                                   //LCom Version V1
                                   #statSend.tsendFct.data[#statSend.tsendFct.dataOffset] := #statSend.configTelegramV1.LComVersion;
                                   #statSend.tsendFct.data[#statSend.tsendFct.dataOffset + 1] := 16#03;
                                   #statSend.tsendFct.data[#statSend.tsendFct.dataOffset + 2] := #statSend.configTelegramV1.comMode;//ComMode
                                   #statSend.tsendFct.data[#statSend.tsendFct.dataOffset + 3] := #statSend.configTelegramV1.slidingWindow;//SlidingWindow
                                   //cycleTime
                                   #statSend.tsendFct.data[#statSend.tsendFct.dataOffset + 4] := #statSend.configTelegramV1.cycleTime.%B1;
                                   #statSend.tsendFct.data[#statSend.tsendFct.dataOffset + 5] := #statSend.configTelegramV1.cycleTime.%B0;
                                   //ackTimeOut
                                   #statSend.tsendFct.data[#statSend.tsendFct.dataOffset + 6] := #statSend.configTelegramV1.ackTimeOut.%B1;
                                   #statSend.tsendFct.data[#statSend.tsendFct.dataOffset + 7] := #statSend.configTelegramV1.ackTimeOut.%B0;
                                   //lifeSignCycle
                                   #statSend.tsendFct.data[#statSend.tsendFct.dataOffset + 8] := #statSend.configTelegramV1.lifeSignCycle.%B1;
                                   #statSend.tsendFct.data[#statSend.tsendFct.dataOffset + 9] := #statSend.configTelegramV1.lifeSignCycle.%B0;
                                   //status
                                   #statSend.tsendFct.data[#statSend.tsendFct.dataOffset + 10] := #statSend.configTelegramV1.status;
                                   //sendModeSyncTime
                                   #statSend.tsendFct.data[#statSend.tsendFct.dataOffset + 11] := #statSend.configTelegramV1.sendModeSyncTime;
                                   //maxSendDataLength
                                   #statSend.tsendFct.data[#statSend.tsendFct.dataOffset + 12] := #statSend.configTelegramV1.maxSendDataLength.%B1;
                                   #statSend.tsendFct.data[#statSend.tsendFct.dataOffset + 13] := #statSend.configTelegramV1.maxSendDataLength.%B0;
                                   //maxReceiveDataLength
                                   #statSend.tsendFct.data[#statSend.tsendFct.dataOffset + 14] := #statSend.configTelegramV1.maxReceiveDataLength.%B1;
                                   #statSend.tsendFct.data[#statSend.tsendFct.dataOffset + 15] := #statSend.configTelegramV1.maxReceiveDataLength.%B0;
                                   //calculate new offset
                                   #statSend.tsendFct.dataOffset := 16;
                               ELSE
                                   #statSend.tsendFct.data[#statSend.tsendFct.dataOffset] := #statSend.configTelegramV2.LComVersion;
                                   #statSend.tsendFct.data[#statSend.tsendFct.dataOffset + 1] := 16#03;
                                   //status
                                   #statSend.tsendFct.data[#statSend.tsendFct.dataOffset + 2] := #statSend.configTelegramV2.status;
                                   //sendModeSyncTime
                                   #statSend.tsendFct.data[#statSend.tsendFct.dataOffset + 3] := #statSend.configTelegramV2.sendModeSyncTime;
                                   //lifeSignCycle
                                   #tempDWord := TIME_TO_DWORD(#statSend.configTelegramV2.lifeSignCycle);
                                   #statSend.tsendFct.data[#statSend.tsendFct.dataOffset + 4] := #tempDWord.%B3;
                                   #statSend.tsendFct.data[#statSend.tsendFct.dataOffset + 5] := #tempDWord.%B2;
                                   #statSend.tsendFct.data[#statSend.tsendFct.dataOffset + 6] := #tempDWord.%B1;
                                   #statSend.tsendFct.data[#statSend.tsendFct.dataOffset + 7] := #tempDWord.%B0;
                                   //cycleTime
                                   #tempDWord := TIME_TO_DWORD(#statSend.configTelegramV2.cycleTime);
                                   #statSend.tsendFct.data[#statSend.tsendFct.dataOffset + 8] := #tempDWord.%B3;
                                   #statSend.tsendFct.data[#statSend.tsendFct.dataOffset + 9] := #tempDWord.%B2;
                                   #statSend.tsendFct.data[#statSend.tsendFct.dataOffset + 10] := #tempDWord.%B1;
                                   #statSend.tsendFct.data[#statSend.tsendFct.dataOffset + 11] := #tempDWord.%B0;
                                   //ackTimeOut
                                   #tempDWord := TIME_TO_DWORD(#statSend.configTelegramV2.ackTimeOut);
                                   #statSend.tsendFct.data[#statSend.tsendFct.dataOffset + 12] := #tempDWord.%B3;
                                   #statSend.tsendFct.data[#statSend.tsendFct.dataOffset + 13] := #tempDWord.%B2;
                                   #statSend.tsendFct.data[#statSend.tsendFct.dataOffset + 14] := #tempDWord.%B1;
                                   #statSend.tsendFct.data[#statSend.tsendFct.dataOffset + 15] := #tempDWord.%B0;
                                   //maxSendDataLength
                                   #statSend.tsendFct.data[#statSend.tsendFct.dataOffset + 16] := #statSend.configTelegramV2.maxSendDataLength.%B3;
                                   #statSend.tsendFct.data[#statSend.tsendFct.dataOffset + 17] := #statSend.configTelegramV2.maxSendDataLength.%B2;
                                   #statSend.tsendFct.data[#statSend.tsendFct.dataOffset + 18] := #statSend.configTelegramV2.maxSendDataLength.%B1;
                                   #statSend.tsendFct.data[#statSend.tsendFct.dataOffset + 19] := #statSend.configTelegramV2.maxSendDataLength.%B0;
                                   //maxReceiveDataLength
                                   #statSend.tsendFct.data[#statSend.tsendFct.dataOffset + 20] := #statSend.configTelegramV2.maxReceiveDataLength.%B3;
                                   #statSend.tsendFct.data[#statSend.tsendFct.dataOffset + 21] := #statSend.configTelegramV2.maxReceiveDataLength.%B2;
                                   #statSend.tsendFct.data[#statSend.tsendFct.dataOffset + 22] := #statSend.configTelegramV2.maxReceiveDataLength.%B1;
                                   #statSend.tsendFct.data[#statSend.tsendFct.dataOffset + 23] := #statSend.configTelegramV2.maxReceiveDataLength.%B0;
                                   //calculate new offset
                                   #statSend.tsendFct.dataOffset := 24;
                               END_IF;
                               #statSend.tsendFct.enable := TRUE;

                               #instLocalLifeSignCycleTimer(IN := FALSE,
                                                            PT := #diagnostics.localConfig.connection.lifeSignCycleTime);
                           ELSE
                               ;//Telegram 3 don´t need be send

                           END_IF;
                       ELSIF (NOT #diagnostics.localConfig.connection.useLComProtocol //without LCom Protocol
                           AND #statState.sender = #STATE_INACTIVE) THEN
                           #statSend.tsendFct.enable := FALSE;
                       ELSE
                           #statSend.tsendFct.enable := TRUE;

                           #instLocalLifeSignCycleTimer(IN := FALSE,
                                                        PT := #diagnostics.localConfig.connection.lifeSignCycleTime);
                       END_IF;

                       //differ between different connection types (IPv4, QDN)
                       IF (#diagnostics.localConfig.connection.connectType = #CON_TYPE_IPV4) THEN
                           #tempConnOucId := #statTconPar.ID;
                       ELSE    //#CON_TYPE_QDN
                           #tempConnOucId := #statTconParQdn.ID;
                       END_IF;

                       #instTSEND(REQ := #statSend.tsendFct.enable,
                                  LEN := #statSend.tsendFct.dataOffset,
                                  ID := #tempConnOucId,
                                  DATA := #statSend.tsendFct.data,
                                  STATUS => #statSend.tsendFct.status);

                       //16#80C4=Temporary communication error
                       IF (#statSend.tsendFct.status = 16#80C4) THEN

                           #instSendErrorTimer(IN := TRUE,
                                               PT := #MAX_TRIAL_TIME);

                           //#MAX_TRIAL_TIME is expired
                           IF #instSendErrorTimer.Q THEN
                               //Write diagnostics
                               #statDiag.bufferIndex := #statDiag.bufferIndex + 1;
                               #statDiag.buffer[#statDiag.bufferIndex].status := #ERR_SEND;
                               #statDiag.buffer[#statDiag.bufferIndex].subFunctionErrorID := #statSend.tsendFct.status;
                               #statDiag.buffer[#statDiag.bufferIndex].additionalValue1 := 0.0;
                               #statDiag.buffer[#statDiag.bufferIndex].additionalValue2 := #statSend.tsendFct.dataOffset;
                               #statDiag.buffer[#statDiag.bufferIndex].additionalValue3 := 0.0;
                               #statDiag.buffer[#statDiag.bufferIndex].additionalValue4 := T#0ms;
                               #statState.connection := #CLOSE_CONNECTION;
                               GOTO diag;
                           END_IF;
                       ELSIF (#statSend.tsendFct.status >= 16#8085) THEN
                           //#WARN_SEND
                           #statDiag.bufferIndex := #statDiag.bufferIndex + 1;
                           #statDiag.buffer[#statDiag.bufferIndex].status := #ERR_SEND;
                           #statDiag.buffer[#statDiag.bufferIndex].subFunctionErrorID := #statSend.tsendFct.status;
                           #statDiag.buffer[#statDiag.bufferIndex].additionalValue1 := 0.0;
                           #statDiag.buffer[#statDiag.bufferIndex].additionalValue2 := #statSend.tsendFct.dataOffset;
                           #statDiag.buffer[#statDiag.bufferIndex].additionalValue3 := 0.0;
                           #statDiag.buffer[#statDiag.bufferIndex].additionalValue4 := T#0ms;

                           #statState.connection := #CLOSE_CONNECTION;
                           GOTO diag;
                       END_IF;
                   END_REGION SEND_LIFESIGN

               END_REGION OPERATION

           #STATE_INACTIVE_PREPARE:
               REGION INACTIVE_PREPARE

                   #statState.connection := #STATE_INACTIVE;
                   #status := #statStatus := #STATUS_NO_CALL;
                   #statFallingEdgeEnable := FALSE;
                   #statOldEnable := FALSE;
                   #busy := FALSE;
               END_REGION INACTIVE_PREPARE

           #STATE_INIT:
               REGION INIT
                   //Reset FB Outputs
                   #connected := #statConnected := FALSE;
                   #sending := #statSending := FALSE;
                   #error := FALSE;

                   //Diagnostics purpose
                   //connection
                   #diagnostics.localConfig.connection.connectionID := #configuration.connection.connectionID;
                   #diagnostics.localConfig.connection.interfaceID := #configuration.connection.interfaceID;
                   #diagnostics.localConfig.connection.comService := #configuration.connection.comService;
                   #diagnostics.localConfig.connection.isClient := #configuration.connection.isClient;
                   #diagnostics.localConfig.connection.localPort := #configuration.connection.localPort;
                   #diagnostics.localConfig.connection.partnerPort := #configuration.connection.partnerPort;
                   #diagnostics.localConfig.connection.partnerIP := #configuration.connection.partnerIP;
                   #diagnostics.localConfig.connection.acceptUnknownPartner := #configuration.connection.acceptUnknownPartner;
                   #statActualLocalLComVersion := #HEADER_V2;
                   #diagnostics.localConfig.connection.lifeSignCycleTime := #configuration.connection.lifeSignCycleTime;
                   //-->QDN
                   #diagnostics.localConfig.connection.connectType := #configuration.connection.connectType;
                   #diagnostics.localConfig.connection.partnerQDN := #configuration.connection.partnerQDN;
                   //Sender
                   #diagnostics.localConfig.sender.cycleTime := #configuration.sender.cycleTime;
                   #diagnostics.localConfig.sender.ackTimeout := #configuration.sender.ackTimeout;
                   //TimeSync
                   #diagnostics.localConfig.timeSync.usePartnerTimestamps := #configuration.timeSync.usePartnerTimestamps;
                   #diagnostics.localConfig.timeSync.sendMode := #configuration.timeSync.sendMode;
                   #diagnostics.localConfig.timeSync.cycleTime := #configuration.timeSync.cycleTime;
                   #diagnostics.localConfig.timeSync.sendAtTimeOfDay := #configuration.timeSync.sendAtTimeOfDay;
                   //Statistics
                   #diagnostics.statistics.avgCallCycle := 0.0;
                   #diagnostics.statistics.avgReceiveMsgCycle := 0.0;
                   #diagnostics.statistics.maxReceiveMsgCycle := T#0ms;
                   #diagnostics.statistics.LComProtocolUsed := FALSE;
                   #diagnostics.statistics.activeLComVersion := 0;
                   #diagnostics.statistics.avgMsgSendingTime := 0.0;
                   #diagnostics.statistics.maxMsgSendingTime := T#0ms;
                   #diagnostics.statistics.avgMsgReceivingTime := 0.0;
                   #diagnostics.statistics.maxMsgReceivingTime := T#0ms;
                   #diagnostics.statistics.numberOfSentMessages := 0;
                   #diagnostics.statistics.numberOfReceivedMessages := 0;
                   #diagnostics.statistics.totalAckTimeouts := 0;
                   #diagnostics.statistics.totalSendCycleViolations := 0;
                   #diagnostics.statistics.totalReceiveCycleViolations := 0;
                   #diagnostics.statistics.totalReconnects := 0;

                   #statConnectAttempts := 0;

                   //Check hardware identifier of the local interface
                   IF ((#diagnostics.localConfig.connection.interfaceID >= 0) //(0...65535)
                       AND
                       (#diagnostics.localConfig.connection.interfaceID <= 65535))
                   THEN
                       //Hardware identifier of the local interface --> OK
                       #statTconPar.InterfaceId := #diagnostics.localConfig.connection.interfaceID;
                   ELSE
                       //Hardware identifier of the local interface --> NOT OK
                       #statDiag.bufferIndex := #statDiag.bufferIndex + 1;
                       #statDiag.buffer[#statDiag.bufferIndex].status := #ERR_INTERFACE_ID;
                       #statDiag.buffer[#statDiag.bufferIndex].subFunctionErrorID := 16#0000;
                       #statDiag.buffer[#statDiag.bufferIndex].additionalValue1 := UINT_TO_REAL(#diagnostics.localConfig.connection.interfaceID);//value from user
                       #statDiag.buffer[#statDiag.bufferIndex].additionalValue2 := 0.0;
                       #statDiag.buffer[#statDiag.bufferIndex].additionalValue3 := 0.0;
                       #statDiag.buffer[#statDiag.bufferIndex].additionalValue4 := T#0ms;

                       #statState.connection := #ERROR_STATE;
                       GOTO diag;
                   END_IF;

                   //Read the IP address
                   #instRDREC(REQ := TRUE,
                              ID := #configuration.connection.interfaceID,
                              INDEX := 16#8080,
                              MLEN := 0,
                              RECORD := #statSend.tsendFct.data);

                   //1st call from RDREC, to get the IP address
                   IF #instRDREC.STATUS = 16#00700100 THEN
                       ;//don´t change the #status = "STATUS_FIRST_CALL"
                   ELSE
                       //change status, that 1st call is just one time occur 
                       #status := #statStatus := #STATUS_INTERMEDIATE_CALL;
                   END_IF;

                   IF (#instRDREC.VALID = TRUE) THEN
                       //New data received and data is valid
                       #diagnostics.localConfig.connection.localIP.ADDR[1] := #statSend.tsendFct.data[28];
                       #diagnostics.localConfig.connection.localIP.ADDR[2] := #statSend.tsendFct.data[29];
                       #diagnostics.localConfig.connection.localIP.ADDR[3] := #statSend.tsendFct.data[30];
                       #diagnostics.localConfig.connection.localIP.ADDR[4] := #statSend.tsendFct.data[31];
                   ELSIF (#instRDREC.ERROR = TRUE) THEN
                       //An error occurred during the reading process
                       #diagnostics.localConfig.connection.localIP.ADDR[1] := 16#00;
                       #diagnostics.localConfig.connection.localIP.ADDR[2] := 16#00;
                       #diagnostics.localConfig.connection.localIP.ADDR[3] := 16#00;
                       #diagnostics.localConfig.connection.localIP.ADDR[4] := 16#00;
                   ELSE
                       RETURN;//The reading process is not complete yet
                   END_IF;

                   //Local port number
                   #statTconPar.LocalPort := #diagnostics.localConfig.connection.localPort;

                   //Check if send buffer is a VARIANT pointer to array of byte
                   IF ((TypeOfElements(#sendBuffer) = TypeOf(#statSend.tsendFct.data[0]))
                       AND
                       (IS_ARRAY(#sendBuffer))) THEN
                       ;//Is VARIANT pointer to array of byte
                   ELSE
                       //Write diagnostics
                       #statDiag.bufferIndex := #statDiag.bufferIndex + 1;
                       #statDiag.buffer[#statDiag.bufferIndex].status := #ERR_SEND_DATA_TYPE;
                       #statDiag.buffer[#statDiag.bufferIndex].subFunctionErrorID := 16#0000;
                       #statDiag.buffer[#statDiag.bufferIndex].additionalValue1 := 0.0;
                       #statDiag.buffer[#statDiag.bufferIndex].additionalValue2 := 0.0;
                       #statDiag.buffer[#statDiag.bufferIndex].additionalValue3 := 0.0;
                       #statDiag.buffer[#statDiag.bufferIndex].additionalValue4 := T#0ms;

                       #statState.connection := #ERROR_STATE;
                       GOTO diag;
                   END_IF;

                   //Check if receive buffer is a VARIANT pointer to array of byte
                   IF ((TypeOfElements(#receiveBuffer) = TypeOf(#statReceive.trcvFct.data[0]))
                       AND
                       (IS_ARRAY(#receiveBuffer))) THEN
                       ;//Is VARIANT pointer to array of byte
                   ELSE
                       //Write diagnostics
                       #statDiag.bufferIndex := #statDiag.bufferIndex + 1;
                       #statDiag.buffer[#statDiag.bufferIndex].status := #ERR_RECEIVE_DATA_TYPE;
                       #statDiag.buffer[#statDiag.bufferIndex].subFunctionErrorID := 16#0000;
                       #statDiag.buffer[#statDiag.bufferIndex].additionalValue1 := 0.0;
                       #statDiag.buffer[#statDiag.bufferIndex].additionalValue2 := 0.0;
                       #statDiag.buffer[#statDiag.bufferIndex].additionalValue3 := 0.0;
                       #statDiag.buffer[#statDiag.bufferIndex].additionalValue4 := T#0ms;

                       #statState.connection := #ERROR_STATE;
                       GOTO diag;
                   END_IF;

                   //Get size of user send buffer and user receive buffer in bytes
                   #diagnostics.localConfig.sizeOfSendBuffer := CountOfElements(#sendBuffer);
                   #diagnostics.localConfig.sizeOfReceiveBuffer := CountOfElements(#receiveBuffer);

                   //Check communication service: 0:UDP, 1:TCP, 2:LCOM
                   IF (#diagnostics.localConfig.connection.comService = 16#01) THEN
                       //Communication service --> transport protocol TCP
                       #statTconPar.ConnectionType := 16#0B;
                       #diagnostics.localConfig.connection.useLComProtocol := FALSE;
                   ELSIF (#diagnostics.localConfig.connection.comService = 16#02) THEN
                       //Communication service --> transport protocol TCP and LCom protocol
                       #statTconPar.ConnectionType := 16#0B;
                       #diagnostics.localConfig.connection.useLComProtocol := TRUE;
                   ELSE
                       //Communication service --> NOT OK
                       //Write diagnostics
                       #statDiag.bufferIndex := #statDiag.bufferIndex + 1;
                       #statDiag.buffer[#statDiag.bufferIndex].status := #ERR_COM_SERVICE;
                       #statDiag.buffer[#statDiag.bufferIndex].subFunctionErrorID := 16#0000;
                       #statDiag.buffer[#statDiag.bufferIndex].additionalValue1 := #diagnostics.localConfig.connection.comService;//value from operator
                       #statDiag.buffer[#statDiag.bufferIndex].additionalValue2 := 0.0;
                       #statDiag.buffer[#statDiag.bufferIndex].additionalValue3 := 0.0;
                       #statDiag.buffer[#statDiag.bufferIndex].additionalValue4 := T#0ms;

                       #statState.connection := #ERROR_STATE;
                       GOTO diag;
                   END_IF;

                   //Check unique connection identifier (16#0001...16#0FFF)
                   IF ((#diagnostics.localConfig.connection.connectionID > 0)
                       AND
                       (#diagnostics.localConfig.connection.connectionID <= 4095))
                   THEN
                       //Connection identifier -->OK
                       #statTconPar.ID := #diagnostics.localConfig.connection.connectionID;
                   ELSE
                       //Connection identifier --> NOT OK
                       //Write diagnostics
                       #statDiag.bufferIndex := #statDiag.bufferIndex + 1;
                       #statDiag.buffer[#statDiag.bufferIndex].status := #ERR_CONNECTION_ID;
                       #statDiag.buffer[#statDiag.bufferIndex].subFunctionErrorID := 16#0000;
                       #statDiag.buffer[#statDiag.bufferIndex].additionalValue1 := WORD_TO_UDINT(#diagnostics.localConfig.connection.connectionID);//value from user
                       #statDiag.buffer[#statDiag.bufferIndex].additionalValue2 := 0.0;
                       #statDiag.buffer[#statDiag.bufferIndex].additionalValue3 := 0.0;
                       #statDiag.buffer[#statDiag.bufferIndex].additionalValue4 := T#0ms;

                       #statState.connection := #ERROR_STATE;
                       GOTO diag;
                   END_IF;

                   //check connection type: 1 = IPv4, 10 = QDN
                   IF (#diagnostics.localConfig.connection.connectType = #CON_TYPE_IPV4) THEN
                       //connection type IPv4
                       ;
                   ELSIF (#diagnostics.localConfig.connection.connectType = #CON_TYPE_QDN) THEN
                       //connection type fully qualified domain name (QDN)
                       ;
                   ELSE
                       //connection type --> NOT OK
                       //write diagnostics
                       #statDiag.bufferIndex := #statDiag.bufferIndex + 1;
                       #statDiag.buffer[#statDiag.bufferIndex].status := #ERR_CONNECTION_TYPE;
                       #statDiag.buffer[#statDiag.bufferIndex].subFunctionErrorID := 16#0000;
                       #statDiag.buffer[#statDiag.bufferIndex].additionalValue1 := #diagnostics.localConfig.connection.connectType;//value from operator
                       #statDiag.buffer[#statDiag.bufferIndex].additionalValue2 := 0.0;
                       #statDiag.buffer[#statDiag.bufferIndex].additionalValue3 := 0.0;
                       #statDiag.buffer[#statDiag.bufferIndex].additionalValue4 := T#0ms;

                       #statState.connection := #ERROR_STATE;
                       GOTO diag;
                   END_IF;

                   //If client
                   IF (#diagnostics.localConfig.connection.isClient) THEN
                       //Partner port and remote address is not checked here
                       //The TCON will rise an error and return value, when the parameters (partnerPort or partnerIP) are wrong
                       //differ between different connection types (IPv4, QDN)
                       IF (#diagnostics.localConfig.connection.connectType = #CON_TYPE_IPV4) THEN
                           //remote addressing via IPv4
                           #statTconPar.RemotePort := #diagnostics.localConfig.connection.partnerPort;
                           #statTconPar.RemoteAddress := #diagnostics.localConfig.connection.partnerIP;
                       ELSE
                           //remote addressing via qualified domain name
                           #statTconParQdn.RemotePort := #diagnostics.localConfig.connection.partnerPort;
                           #statTconParQdn.RemoteQDN := #diagnostics.localConfig.connection.partnerQDN;
                           //additionally store all TCON configurations done before for QDN connection parameters
                           #statTconParQdn.ConnectionType := 16#0B;
                           #statTconParQdn.LocalPort := #diagnostics.localConfig.connection.localPort;
                           #statTconParQdn.InterfaceId := #diagnostics.localConfig.connection.interfaceID;
                           #statTconParQdn.ID := #diagnostics.localConfig.connection.connectionID;
                       END_IF;
                       //If server
                   ELSE
                       //Accept requests from all partners or only specified partner is allowed
                       IF (#diagnostics.localConfig.connection.acceptUnknownPartner) THEN
                           //Accept requests from all partners
                           //differ between different connection types (IPv4, QDN)
                           IF (#diagnostics.localConfig.connection.connectType = #CON_TYPE_IPV4) THEN
                               #statTconPar.RemoteAddress.ADDR[1] := 0;
                               #statTconPar.RemoteAddress.ADDR[2] := 0;
                               #statTconPar.RemoteAddress.ADDR[3] := 0;
                               #statTconPar.RemoteAddress.ADDR[4] := 0;
                               #statTconPar.RemotePort := 0;
                           ELSE    //#CON_TYPE_QDN
                               #statTconParQdn.RemoteQDN := '';
                               #statTconParQdn.RemotePort := 0;
                           END_IF;
                       ELSE
                           //Only specified partner is allowed
                           //differ between different connection types (IPv4, QDN)
                           IF (#diagnostics.localConfig.connection.connectType = #CON_TYPE_IPV4) THEN
                               #statTconPar.RemoteAddress := #diagnostics.localConfig.connection.partnerIP;
                               #statTconPar.RemotePort := #diagnostics.localConfig.connection.partnerPort;
                           ELSE    //#CON_TYPE_QDN
                               #statTconParQdn.RemoteQDN := #diagnostics.localConfig.connection.partnerQDN;
                               #statTconParQdn.RemotePort := #diagnostics.localConfig.connection.partnerPort;
                           END_IF;
                       END_IF;
                   END_IF;

                   //Check cycleTime
                   IF ((#diagnostics.localConfig.sender.cycleTime >= T#0ms)
                       AND
                       (#diagnostics.localConfig.sender.cycleTime <= T#+24d20h31m23s647ms))
                   THEN
                       ;//CycleTime --> OK
                   ELSE
                       //CycleTime --> NOT OK
                       #statDiag.bufferIndex := #statDiag.bufferIndex + 1;
                       #statDiag.buffer[#statDiag.bufferIndex].status := #ERR_SEND_CYCLE_TIME;
                       #statDiag.buffer[#statDiag.bufferIndex].subFunctionErrorID := 16#0000;
                       #statDiag.buffer[#statDiag.bufferIndex].additionalValue1 := 0.0;
                       #statDiag.buffer[#statDiag.bufferIndex].additionalValue2 := 0.0;
                       #statDiag.buffer[#statDiag.bufferIndex].additionalValue3 := 0.0;
                       #statDiag.buffer[#statDiag.bufferIndex].additionalValue4 := #diagnostics.localConfig.sender.cycleTime;//value from operator

                       #statState.connection := #ERROR_STATE;
                       GOTO diag;
                   END_IF;

                   //With LCom header
                   IF (#diagnostics.localConfig.connection.useLComProtocol) THEN

                       //Check lifeSignCycleTime
                       IF ((#diagnostics.localConfig.connection.lifeSignCycleTime > T#0ms) //(1ms...T#+24d20h31m23s647ms)
                           AND
                           (#diagnostics.localConfig.connection.lifeSignCycleTime <= T#+24d20h31m23s647ms))
                       THEN
                           ;//lifeSignCycleTime--> OK
                       ELSE
                           //LifeSignCycle --> NOT OK
                           #statDiag.bufferIndex := #statDiag.bufferIndex + 1;
                           #statDiag.buffer[#statDiag.bufferIndex].status := #ERR_LIFE_SIGN_CYCLE;
                           #statDiag.buffer[#statDiag.bufferIndex].subFunctionErrorID := 16#0000;
                           #statDiag.buffer[#statDiag.bufferIndex].additionalValue1 := 0.0;
                           #statDiag.buffer[#statDiag.bufferIndex].additionalValue2 := 0.0;
                           #statDiag.buffer[#statDiag.bufferIndex].additionalValue3 := 0.0;
                           #statDiag.buffer[#statDiag.bufferIndex].additionalValue4 := #diagnostics.localConfig.connection.lifeSignCycleTime;//value from operator

                           #statState.connection := #ERROR_STATE;
                           GOTO diag;
                       END_IF;

                       //Check ackTimeOut
                       IF ((#diagnostics.localConfig.sender.ackTimeout > T#0ms)
                           AND
                           (#diagnostics.localConfig.sender.ackTimeout <= T#+24d20h31m23s647ms))
                       THEN
                           ;//AckTimeOut --> OK
                       ELSE
                           //AckTimeOut --> NOT OK
                           #statDiag.bufferIndex := #statDiag.bufferIndex + 1;
                           #statDiag.buffer[#statDiag.bufferIndex].status := #ERR_ACK_TIMEOUT;
                           #statDiag.buffer[#statDiag.bufferIndex].subFunctionErrorID := 16#0000;
                           #statDiag.buffer[#statDiag.bufferIndex].additionalValue1 := 0.0;
                           #statDiag.buffer[#statDiag.bufferIndex].additionalValue2 := 0.0;
                           #statDiag.buffer[#statDiag.bufferIndex].additionalValue3 := 0.0;
                           #statDiag.buffer[#statDiag.bufferIndex].additionalValue4 := #diagnostics.localConfig.sender.ackTimeout;//value from operator

                           #statState.connection := #ERROR_STATE;
                           GOTO diag;
                       END_IF;

                       //Check timeSync
                       IF (NOT #diagnostics.localConfig.timeSync.usePartnerTimestamps) THEN

                           IF ((#diagnostics.localConfig.timeSync.sendMode >= 0)//(0...2)
                               AND
                               (#diagnostics.localConfig.timeSync.sendMode <= 2))
                           THEN
                               CASE (#diagnostics.localConfig.timeSync.sendMode) OF

                                   1: //TimeSync.cycleTime
                                       IF ((#diagnostics.localConfig.timeSync.cycleTime > T#0ms) //(1ms...T#+24d20h31m23s647ms)
                                           AND
                                           (#diagnostics.localConfig.timeSync.cycleTime <= T#+24d20h31m23s647ms))
                                       THEN
                                           ;//CycleTime --> OK
                                       ELSE
                                           //CycleTime --> Not OK
                                           #statDiag.bufferIndex := #statDiag.bufferIndex + 1;
                                           #statDiag.buffer[#statDiag.bufferIndex].status := #ERR_TIME_CYCLE_TIME;
                                           #statDiag.buffer[#statDiag.bufferIndex].subFunctionErrorID := 16#0000;
                                           #statDiag.buffer[#statDiag.bufferIndex].additionalValue1 := 0.0;
                                           #statDiag.buffer[#statDiag.bufferIndex].additionalValue2 := 0.0;
                                           #statDiag.buffer[#statDiag.bufferIndex].additionalValue3 := 0.0;
                                           #statDiag.buffer[#statDiag.bufferIndex].additionalValue4 := #diagnostics.localConfig.timeSync.cycleTime;//value from user

                                           #statState.connection := #ERROR_STATE;
                                           GOTO diag;

                                       END_IF;
                                   2://TimeSync.sendAtTimeOfDay
                                       IF ((#diagnostics.localConfig.timeSync.sendAtTimeOfDay >= TOD#00:00:00.000) //(TOD#00:00:00.000...TOD#23:59:59.999)
                                           AND
                                           #diagnostics.localConfig.timeSync.sendAtTimeOfDay <= TOD#23:59:59.999)
                                       THEN
                                           ;//SendAtTimeOfDay --> OK
                                       ELSE
                                           //SendAtTimeOfDay --> NOT OK
                                           #statDiag.bufferIndex := #statDiag.bufferIndex + 1;
                                           #statDiag.buffer[#statDiag.bufferIndex].status := #ERR_TIME_OF_DAY;
                                           #statDiag.buffer[#statDiag.bufferIndex].subFunctionErrorID := 16#0000;
                                           #statDiag.buffer[#statDiag.bufferIndex].additionalValue1 := 0.0;
                                           #statDiag.buffer[#statDiag.bufferIndex].additionalValue2 := 0.0;
                                           #statDiag.buffer[#statDiag.bufferIndex].additionalValue3 := 0.0;
                                           #statDiag.buffer[#statDiag.bufferIndex].additionalValue4 := T#0ms;

                                           #statState.connection := #ERROR_STATE;
                                           GOTO diag;
                                       END_IF;
                                   ELSE
                                       ;
                               END_CASE;
                           ELSE
                               //SendMode --> NOT OK
                               #statDiag.bufferIndex := #statDiag.bufferIndex + 1;
                               #statDiag.buffer[#statDiag.bufferIndex].status := #ERR_TIME_SYNC_MODE;
                               #statDiag.buffer[#statDiag.bufferIndex].subFunctionErrorID := 16#0000;
                               #statDiag.buffer[#statDiag.bufferIndex].additionalValue1 := #diagnostics.localConfig.timeSync.sendMode;
                               #statDiag.buffer[#statDiag.bufferIndex].additionalValue2 := 0.0;
                               #statDiag.buffer[#statDiag.bufferIndex].additionalValue3 := 0.0;
                               #statDiag.buffer[#statDiag.bufferIndex].additionalValue4 := T#0ms;

                               #statState.connection := #ERROR_STATE;
                               GOTO diag;
                           END_IF;
                       ELSE
                           //usePartnerTimeStamp

                           //Is sendMode inactive ?
                           IF #diagnostics.localConfig.timeSync.sendMode = 0 THEN
                               ;// Yes
                           ELSE
                               //SendMode --> NOT OK
                               #statDiag.bufferIndex := #statDiag.bufferIndex + 1;
                               #statDiag.buffer[#statDiag.bufferIndex].status := #ERR_TIME_SYNC_MODE;
                               #statDiag.buffer[#statDiag.bufferIndex].subFunctionErrorID := 16#0000;
                               #statDiag.buffer[#statDiag.bufferIndex].additionalValue1 := #diagnostics.localConfig.timeSync.sendMode;
                               #statDiag.buffer[#statDiag.bufferIndex].additionalValue2 := 0.0;
                               #statDiag.buffer[#statDiag.bufferIndex].additionalValue3 := 0.0;
                               #statDiag.buffer[#statDiag.bufferIndex].additionalValue4 := T#0ms;

                               #statState.connection := #ERROR_STATE;
                               GOTO diag;
                           END_IF;

                       END_IF;
                   ELSE
                       ;//No LCom Protocol is used
                   END_IF;

                   //differ between different connection types (IPv4, QDN)
                   IF (#diagnostics.localConfig.connection.connectType = #CON_TYPE_IPV4) THEN
                       //IPv4
                       #instTCON(REQ := FALSE,
                                 ID := #statTconPar.ID,
                                 CONNECT := #statTconPar);
                       //store connection ID temporary
                       #tempConnOucId := #statTconPar.ID;
                   ELSE
                       //QDN (CON_TYPE_QDN)
                       #instTCON(REQ := FALSE,
                                 ID := #statTconParQdn.ID,
                                 CONNECT := #statTconParQdn);
                       //store connection ID temporary
                       #tempConnOucId := #statTconParQdn.ID;
                   END_IF;

                   #instTSEND(REQ := FALSE,
                              ID := #tempConnOucId,
                              DATA := #statSend.tsendFct.data);

                   #instTRCV(EN_R := FALSE,
                             ID := #tempConnOucId,
                             DATA := #statReceive.trcvFct.data);

                   #instTDISCON(REQ := FALSE,
                                ID := #tempConnOucId);

                   //Passive (server), active connection establishment (client)
                   IF (#diagnostics.localConfig.connection.isClient) THEN
                       #statState.connection := #OPEN_CLIENT;
                       #statTconPar.ActiveEstablished := TRUE;
                       #statTconParQdn.ActiveEstablished := TRUE;
                   ELSE
                       #statState.connection := #OPEN_SERVER;
                       #statTconPar.ActiveEstablished := FALSE;
                       #statTconParQdn.ActiveEstablished := FALSE;
                   END_IF;
               END_REGION INIT

           #OPEN_CLIENT, #OPEN_SERVER:
               REGION OPEN_CLIENT_SERVER
                   #instTCON.STATUS := 16#0000;

                   //differ between different connection types (IPv4, QDN)
                   IF (#diagnostics.localConfig.connection.connectType = #CON_TYPE_IPV4) THEN
                       //IPv4
                       #instTCON(REQ := TRUE,
                                 CONNECT := #statTconPar,
                                 ID := #diagnostics.localConfig.connection.connectionID);
                   ELSE
                       //QDN (CON_TYPE_QDN)
                       #instTCON(REQ := TRUE,
                                 CONNECT := #statTconParQdn,
                                 ID := #diagnostics.localConfig.connection.connectionID);
                   END_IF;

                   // Error occurred
                   IF (#instTCON.ERROR) THEN

                       //Local port is being used by the system
                       IF (#instTCON.STATUS = 16#80A2 OR (#diagnostics.localConfig.connection.connectType = #CON_TYPE_IPV4 AND #statTconPar.LocalPort = 16#0)) THEN

                           #statDiag.bufferIndex := #statDiag.bufferIndex + 1;
                           #statDiag.buffer[#statDiag.bufferIndex].status := #ERR_LOCAL_PORT;
                           #statDiag.buffer[#statDiag.bufferIndex].subFunctionErrorID := #instTCON.STATUS;
                           #statDiag.buffer[#statDiag.bufferIndex].additionalValue1 := #statTconPar.LocalPort;
                           #statDiag.buffer[#statDiag.bufferIndex].additionalValue2 := 0.0;
                           #statDiag.buffer[#statDiag.bufferIndex].additionalValue3 := 0.0;
                           #statDiag.buffer[#statDiag.bufferIndex].additionalValue4 := T#0ms;

                           #statState.connection := #ERROR_STATE;
                           GOTO diag;
                           //Local port is being used by the system (in case of QDN)
                       ELSIF (#instTCON.STATUS = 16#80A2 OR (#diagnostics.localConfig.connection.connectType = #CON_TYPE_QDN AND #statTconParQdn.LocalPort = 16#0)) THEN

                           #statDiag.bufferIndex := #statDiag.bufferIndex + 1;
                           #statDiag.buffer[#statDiag.bufferIndex].status := #ERR_LOCAL_PORT;
                           #statDiag.buffer[#statDiag.bufferIndex].subFunctionErrorID := #instTCON.STATUS;
                           #statDiag.buffer[#statDiag.bufferIndex].additionalValue1 := #statTconParQdn.LocalPort;
                           #statDiag.buffer[#statDiag.bufferIndex].additionalValue2 := 0.0;
                           #statDiag.buffer[#statDiag.bufferIndex].additionalValue3 := 0.0;
                           #statDiag.buffer[#statDiag.bufferIndex].additionalValue4 := T#0ms;

                           #statState.connection := #ERROR_STATE;
                           GOTO diag;
                       ELSIF (#instTCON.STATUS = 16#80B7 OR #instTCON.STATUS = 16#80A4) THEN
                           //IP address of the remote partner is invalid
                           #statDiag.bufferIndex := #statDiag.bufferIndex + 1;
                           #statDiag.buffer[#statDiag.bufferIndex].status := #ERR_PARTNER_IP;
                           #statDiag.buffer[#statDiag.bufferIndex].subFunctionErrorID := #instTCON.STATUS;
                           #statDiag.buffer[#statDiag.bufferIndex].additionalValue1 := 0.0;
                           #statDiag.buffer[#statDiag.bufferIndex].additionalValue2 := 0.0;
                           #statDiag.buffer[#statDiag.bufferIndex].additionalValue3 := 0.0;
                           #statDiag.buffer[#statDiag.bufferIndex].additionalValue4 := T#0ms;

                           #statState.connection := #ERROR_STATE;
                           GOTO diag;
                       ELSIF (#instTCON.STATUS = 16#809B) THEN
                           //The local_device_id in the connection description does not match the CPU
                           #statDiag.bufferIndex := #statDiag.bufferIndex + 1;
                           #statDiag.buffer[#statDiag.bufferIndex].status := #ERR_INTERFACE_ID;
                           #statDiag.buffer[#statDiag.bufferIndex].subFunctionErrorID := #instTCON.STATUS;
                           #statDiag.buffer[#statDiag.bufferIndex].additionalValue1 := UINT_TO_REAL(#diagnostics.localConfig.connection.interfaceID);//value from user
                           #statDiag.buffer[#statDiag.bufferIndex].additionalValue2 := 0.0;
                           #statDiag.buffer[#statDiag.bufferIndex].additionalValue3 := 0.0;
                           #statDiag.buffer[#statDiag.bufferIndex].additionalValue4 := T#0ms;

                           #statState.connection := #ERROR_STATE;
                           GOTO diag;
                       ELSE
                           IF (#statState.connection = #OPEN_CLIENT) THEN

                               #statDiag.bufferIndex := #statDiag.bufferIndex + 1;
                               #statDiag.buffer[#statDiag.bufferIndex].status := #ERR_OPEN_CLIENT;
                               #statDiag.buffer[#statDiag.bufferIndex].subFunctionErrorID := #instTCON.STATUS;
                               #statDiag.buffer[#statDiag.bufferIndex].additionalValue1 := 0.0;
                               #statDiag.buffer[#statDiag.bufferIndex].additionalValue2 := 0.0;
                               #statDiag.buffer[#statDiag.bufferIndex].additionalValue3 := 0.0;
                               #statDiag.buffer[#statDiag.bufferIndex].additionalValue4 := T#0ms;

                               //Try reconnection after a wait time
                               #statIterator := 0;
                               #statState.connection := #STATE_WAIT;
                           ELSE
                               #statDiag.bufferIndex := #statDiag.bufferIndex + 1;
                               #statDiag.buffer[#statDiag.bufferIndex].status := #ERR_OPEN_SERVER;
                               #statDiag.buffer[#statDiag.bufferIndex].subFunctionErrorID := #instTCON.STATUS;
                               //differ between different connection types (IPv4, QDN)
                               IF (#diagnostics.localConfig.connection.connectType = #CON_TYPE_IPV4) THEN
                                   #statDiag.buffer[#statDiag.bufferIndex].additionalValue1 := #statTconPar.LocalPort;
                               ELSE    //CON_TYPE_QDN
                                   #statDiag.buffer[#statDiag.bufferIndex].additionalValue1 := #statTconParQdn.LocalPort;
                               END_IF;
                               #statDiag.buffer[#statDiag.bufferIndex].additionalValue2 := 0.0;
                               #statDiag.buffer[#statDiag.bufferIndex].additionalValue3 := 0.0;
                               #statDiag.buffer[#statDiag.bufferIndex].additionalValue4 := T#0ms;

                               //Try reconnection after a wait time
                               #statIterator := 0;
                               #statState.connection := #STATE_WAIT;
                           END_IF;
                       END_IF;
                       //Job completed without error
                   ELSIF (#instTCON.DONE) THEN

                       //Connection successfully established
                       #diagnostics.statistics.totalReconnects := #diagnostics.statistics.totalReconnects + 1;
                       #statState.connection := #OPERATION;

                       #error := FALSE;

                       //Reset all state machines
                       #statState.receiver := #READ;
                       #statState.sender := #STATE_INACTIVE;
                       #statState.comReceiver := #EXPECTED;
                       #statState.comSender := #STATE_INACTIVE;
                       //Receive
                       #statReceive.trcvFct.dataOffset := 0;
                       #statReceive.trcvFct.dataLength := 0;
                       #statReceive.trcvFct.dataLengthRest := 0;
                       #statReceive.trcvFct.dataReceived := FALSE;
                       #statReceive.tempTelegram.index := 0;
                       #statReceive.tempTelegram.telegramType := 0;
                       #statReceive.numberOfLComHeader := 0;
                       #statReceive.dataTelegram.totalMessageLength := 0;
                       #statReceive.dataTelegram.actPackageLength := 0;
                       #statReceive.dataTelegram.ackMessageOffset := 0;
                       #statReceive.dataTelegram.messageOffset := 0;
                       #statReceive.dataTelegram.ackMessageCounter := 0;
                       #statReceive.dataTelegram.messageCounter := 0;
                       #statReceive.userData.totalLength := 0;
                       #statReceive.userData.offset := 0;
                       //Send
                       #statSend.tsendFct.dataLengthRest := 0;
                       #statSend.tsendFct.dataOffset := 0;
                       #statSend.tsendFct.status := 16#0000;
                       #statSend.expectedAck.package1.offset := 0;
                       #statSend.dataTelegram.messageCounter := 0;
                       #statSend.dataTelegram.ackMessageCounter := 0;
                       #statSend.dataTelegram.messageOffset := 0;
                       #statSend.dataTelegram.ackMessageOffset := 0;
                       #statSend.dataTelegram.actPackageLength := 0;
                       #statSend.dataTelegram.totalMessageLength := 0;
                       #statSend.numberOfLComPackage := 0;
                       #statSend.userData.totalLength := 0;
                       #statSend.userData.offset := 0;
                       #statSend.userData.sendCycleViolation := FALSE;
                       #statOldSend := FALSE;

                       #diagnostics.statistics.maxMsgSendingTime := T#0ms;
                       #diagnostics.localConfig.sender.cycleTime := T#0ms;
                       #diagnostics.localConfig.sender.ackTimeout := T#0ms;

                       #diagnostics.statistics.lastTimeSync.YEAR := 2200;
                       #statCopyNBytes := 0;

                       //Reset all timer
                       #instLocalLifeSignCycleTimer(IN := FALSE,
                                                    PT := #diagnostics.localConfig.connection.lifeSignCycleTime);

                       #instPartnerLifeSignCycleTimer(IN := FALSE,
                                                      PT := (#diagnostics.partnerConfig.connnection.lifeSignCycleTime));

                       #instLocalCycleTimeTimer(IN := FALSE,
                                                PT := #diagnostics.localConfig.sender.cycleTime);

                       #instExpectedAckPackage1(IN := FALSE,
                                                PT := #diagnostics.localConfig.sender.ackTimeout);

                       #instSyncTimer(IN := FALSE,
                                      PT := T#1s);

                       #instSendErrorTimer(IN := FALSE,
                                           PT := #MAX_TRIAL_TIME);

                       #instRcvErrorTimer(IN := FALSE,
                                          PT := #MAX_TRIAL_TIME);

                       //Reset all active failures in the diagnostics buffer
                       FOR #statIterator := 0 TO #DIAG_BUFFER_UPPER_LIM BY 1 DO
                           #diagnostics.buffer[#statIterator].isActive := FALSE;
                       END_FOR;

                       //With LCom protocol
                       IF (#diagnostics.localConfig.connection.useLComProtocol = TRUE) THEN

                           IF (#statConnectAttempts MOD 2 = 0) THEN
                               //1st try LCom Version 2.0
                               #statActualLocalLComVersion := #HEADER_V2;
                               #statSend.configTelegramV2.LComVersion := #HEADER_V2;
                               #statSend.configTelegramV2.status := BOOL_TO_BYTE(#diagnostics.localConfig.timeSync.usePartnerTimestamps);
                               #statSend.configTelegramV2.sendModeSyncTime := #diagnostics.localConfig.timeSync.sendMode;
                               #statSend.configTelegramV2.lifeSignCycle := #diagnostics.localConfig.connection.lifeSignCycleTime;
                               #statSend.configTelegramV2.cycleTime := #configuration.sender.cycleTime;
                               #statSend.configTelegramV2.ackTimeOut := #configuration.sender.ackTimeout;
                               #statSend.configTelegramV2.maxSendDataLength := #diagnostics.localConfig.sizeOfSendBuffer;
                               #statSend.configTelegramV2.maxReceiveDataLength := #diagnostics.localConfig.sizeOfReceiveBuffer;

                               #statSend.dataTelegram.LComVersion := #statSend.configTelegramV2.LComVersion;
                           ELSE
                               //2nd try LCom Version 1.0
                               #statActualLocalLComVersion := #HEADER_V1;
                               #statSend.configTelegramV1.LComVersion := #HEADER_V1;
                               #statSend.configTelegramV1.comMode := 16#03;
                               #statSend.configTelegramV1.slidingWindow := 1;
                               #statSend.configTelegramV1.status := BOOL_TO_BYTE(#diagnostics.localConfig.timeSync.usePartnerTimestamps);
                               #statSend.configTelegramV1.sendModeSyncTime := #diagnostics.localConfig.timeSync.sendMode;

                               #statSend.dataTelegram.LComVersion := #statSend.configTelegramV1.LComVersion;

                               //Check max. lifeSignCycleTime
                               IF (#diagnostics.localConfig.connection.lifeSignCycleTime > T#65535ms) THEN

                                   #statDiag.bufferIndex := #statDiag.bufferIndex + 1;
                                   #statDiag.buffer[#statDiag.bufferIndex].additionalValue4 := #diagnostics.localConfig.connection.lifeSignCycleTime;
                                   #diagnostics.localConfig.connection.lifeSignCycleTime := T#65535ms;

                                   #statDiag.buffer[#statDiag.bufferIndex].status := #WARN_LIFE_SIGN_LIMITATION;
                                   #statDiag.buffer[#statDiag.bufferIndex].subFunctionErrorID := 16#0000;
                                   #statDiag.buffer[#statDiag.bufferIndex].additionalValue1 := 65535.0;
                                   #statDiag.buffer[#statDiag.bufferIndex].additionalValue2 := 0.0;
                                   #statDiag.buffer[#statDiag.bufferIndex].additionalValue3 := 0.0;
                               ELSE
                                   ;
                               END_IF;
                               #statSend.configTelegramV1.lifeSignCycle := TIME_TO_UINT(#diagnostics.localConfig.connection.lifeSignCycleTime);

                               //Check max.sizeOfSendBuffer
                               IF (#diagnostics.localConfig.sizeOfSendBuffer > 65535) THEN
                                   #diagnostics.localConfig.sizeOfSendBuffer := 65535;
                                   #statSend.configTelegramV1.maxSendDataLength := 65535;
                               ELSE
                                   #statSend.configTelegramV1.maxSendDataLength := UDINT_TO_UINT(#diagnostics.localConfig.sizeOfSendBuffer);
                               END_IF;

                               //Check max.sizeOfReceiveBuffer
                               IF (#diagnostics.localConfig.sizeOfReceiveBuffer > 65535) THEN
                                   #diagnostics.localConfig.sizeOfReceiveBuffer := 65535;
                                   #statSend.configTelegramV1.maxReceiveDataLength := 65535;
                               ELSE
                                   #statSend.configTelegramV1.maxReceiveDataLength := UDINT_TO_UINT(#diagnostics.localConfig.sizeOfReceiveBuffer);
                               END_IF;

                           END_IF;
                           //Set telegram type of data telegrams for LCom Version 1.0 and 2.0
                           #statSend.dataTelegram.telegramType := 16#0A;

                           //Start sender config directly with LCom protocol
                           #statState.cfgSender := #STATE_INIT;
                       ELSE
                           //without LCom
                           #statCompare.sender.cycleTime := #configuration.sender.cycleTime;
                           #diagnostics.localConfig.sender.cycleTime := #configuration.sender.cycleTime;

                           #diagnostics.partnerConfig.sizeOfReceiveBuffer := 0;
                           #diagnostics.partnerConfig.sizeOfSendBuffer := 0;
                           #connected := #statConnected := TRUE;
                           #statState.cfgSender := #OPERATION;

                           #statDiag.bufferIndex := #statDiag.bufferIndex + 1;
                           #statDiag.buffer[#statDiag.bufferIndex].status := #STATUS_TCP_CONNECTED;
                           #statDiag.buffer[#statDiag.bufferIndex].subFunctionErrorID := 16#0000;
                           #statDiag.buffer[#statDiag.bufferIndex].additionalValue1 := 0.0;
                           #statDiag.buffer[#statDiag.bufferIndex].additionalValue2 := 0.0;
                           #statDiag.buffer[#statDiag.bufferIndex].additionalValue3 := 0.0;
                           #statDiag.buffer[#statDiag.bufferIndex].additionalValue4 := T#0ms;
                       END_IF;
                       //TCON still in progress
                   ELSE
                       IF (#diagnostics.localConfig.connection.isClient) THEN

                           #statDiag.bufferIndex := #statDiag.bufferIndex + 1;
                           #statDiag.buffer[#statDiag.bufferIndex].status := #STATUS_CLIENT_TRY_CONNECT;
                           #statDiag.buffer[#statDiag.bufferIndex].subFunctionErrorID := 16#0000;
                           #statDiag.buffer[#statDiag.bufferIndex].additionalValue1 := 0.0;
                           #statDiag.buffer[#statDiag.bufferIndex].additionalValue2 := 0.0;
                           #statDiag.buffer[#statDiag.bufferIndex].additionalValue3 := 0.0;
                           #statDiag.buffer[#statDiag.bufferIndex].additionalValue4 := T#0ms;
                       ELSE
                           #statDiag.bufferIndex := #statDiag.bufferIndex + 1;
                           #statDiag.buffer[#statDiag.bufferIndex].status := #STATUS_SERVER_PORT_OPEN;
                           #statDiag.buffer[#statDiag.bufferIndex].subFunctionErrorID := 16#0000;
                           #statDiag.buffer[#statDiag.bufferIndex].additionalValue1 := 0.0;
                           #statDiag.buffer[#statDiag.bufferIndex].additionalValue2 := 0.0;
                           #statDiag.buffer[#statDiag.bufferIndex].additionalValue3 := 0.0;
                           #statDiag.buffer[#statDiag.bufferIndex].additionalValue4 := T#0ms;
                       END_IF;
                   END_IF;
               END_REGION OPEN_CLIENT_SERVER

           #STATE_WAIT:
               REGION WAIT
                   //Wait and then establish the connection
                   IF (#statIterator > #STATE_WAIT) THEN

                       #tempConnOucId := 0;

                       //differ between different connection types (IPv4, QDN)
                       IF (#diagnostics.localConfig.connection.connectType = #CON_TYPE_IPV4) THEN
                           //IPv4
                           #instTCON(REQ := FALSE,
                                     ID := #statTconPar.ID,
                                     CONNECT := #statTconPar);
                           //store connection ID temporary
                           #tempConnOucId := #statTconPar.ID;
                       ELSE
                           //QDN (CON_TYPE_QDN)
                           #instTCON(REQ := FALSE,
                                     ID := #statTconParQdn.ID,
                                     CONNECT := #statTconParQdn);
                           //store connection ID temporary
                           #tempConnOucId := #statTconParQdn.ID;
                       END_IF;

                       #instTSEND(REQ := FALSE,
                                  ID := #tempConnOucId,
                                  DATA := #statSend.tsendFct.data);

                       #instTRCV(EN_R := FALSE,
                                 ID := #tempConnOucId,
                                 DATA := #statReceive.trcvFct.data);

                       #instTDISCON(REQ := FALSE,
                                    ID := #tempConnOucId);

                       IF (#diagnostics.localConfig.connection.isClient) THEN
                           #statState.connection := #OPEN_CLIENT;
                           #statTconPar.ActiveEstablished := TRUE;
                           #statTconParQdn.ActiveEstablished := TRUE;
                       ELSE
                           #statState.connection := #OPEN_SERVER;
                           #statTconPar.ActiveEstablished := FALSE;
                           #statTconParQdn.ActiveEstablished := FALSE;
                       END_IF;

                   ELSE
                       #statIterator := #statIterator + 1;
                   END_IF;
               END_REGION WAIT

           #FINISH_TSEND:
               REGION FINISH_TSEND
                   IF (#statIterator > #STATE_WAIT) THEN
                       #statIterator := 0;
                       #statState.connection := #FINISH_TRCV;
                   ELSE
                       //differ between different connection types (IPv4, QDN)
                       IF (#diagnostics.localConfig.connection.connectType = #CON_TYPE_IPV4) THEN
                           #tempConnOucId := #statTconPar.ID;
                       ELSE    //CON_TYPE_QDN
                           #tempConnOucId := #statTconParQdn.ID;
                       END_IF;

                       #instTSEND(REQ := TRUE,
                                  LEN := #statSend.tsendFct.dataOffset,
                                  ID := #tempConnOucId,
                                  DATA := #statSend.tsendFct.data,
                                  STATUS => #statSend.tsendFct.status);

                       IF ((#statSend.tsendFct.status = 16#0000) OR (#instTSEND.ERROR)) THEN
                           //"TSEND" instruction is finished
                           #statState.connection := #FINISH_TRCV;
                       ELSE
                           ;//"TSEND" instruction still in process
                       END_IF;
                   END_IF;
                   #statIterator := #statIterator + 1;
               END_REGION FINISH_TSEND

           #FINISH_TRCV:
               REGION FINISH_TRCV

                   IF (#statIterator > #STATE_WAIT) THEN
                       #statState.connection := #CALL_TDISCON;
                   ELSE
                       //differ between different connection types (IPv4, QDN)
                       IF (#diagnostics.localConfig.connection.connectType = #CON_TYPE_IPV4) THEN
                           #tempConnOucId := #statTconPar.ID;
                       ELSE    //CON_TYPE_QDN
                           #tempConnOucId := #statTconParQdn.ID;
                       END_IF;

                       #instTRCV(EN_R := TRUE,
                                 ID := #tempConnOucId,
                                 LEN := 0,
                                 ADHOC := TRUE,
                                 NDR => #statReceive.trcvFct.dataReceived,
                                 RCVD_LEN => #statReceive.trcvFct.dataLength,
                                 DATA := #statReceive.trcvFct.data);

                       //Is the "TRCV" instruction still in process
                       IF (#instTRCV.ERROR OR NOT #instTRCV.BUSY) THEN
                           #statState.connection := #CALL_TDISCON;
                       ELSE
                           ;//TRCV instruction still in process
                       END_IF;
                   END_IF;
                   #statIterator := #statIterator + 1;
               END_REGION FINISH_TRCV

           #CLOSE_CONNECTION:
               REGION CLOSE_CONNECTION
                   //reset FB Outputs
                   #connected := #statConnected := FALSE;
                   #sending := #statSending := FALSE;
                   #receivedDataLength := 0;
                   #error := FALSE;

                   //Is "TSEND" instruction still in process ?
                   IF (#statSend.tsendFct.status <> 16#0000) THEN
                       //"TSEND" instruction still in process
                       #statState.connection := #FINISH_TSEND;
                       #statIterator := 0;
                   ELSE
                       ;//"TSEND" instruction is finished
                   END_IF;

                   #instTRCV(EN_R := TRUE,
                             ID := #diagnostics.localConfig.connection.connectionID,
                             LEN := 0,
                             ADHOC := TRUE,
                             NDR => #statReceive.trcvFct.dataReceived,
                             RCVD_LEN => #statReceive.trcvFct.dataLength,
                             DATA := #statReceive.trcvFct.data);

                   //Is the "TRCV" instruction still in process
                   IF (#instTRCV.ERROR OR NOT #instTRCV.BUSY) THEN
                       #statState.connection := #CALL_TDISCON;
                   ELSE
                       #statState.connection := #FINISH_TRCV;
                       #statIterator := 0;
                   END_IF;
               END_REGION CLOSE_CONNECTION

           #CALL_TDISCON:
               REGION CALL_TDISCON
                   //differ between different connection types (IPv4, QDN)
                   IF (#diagnostics.localConfig.connection.connectType = #CON_TYPE_IPV4) THEN
                       #tempConnOucId := #statTconPar.ID;
                   ELSE    //CON_TYPE_QDN
                       #tempConnOucId := #statTconParQdn.ID;
                   END_IF;

                   #instTSEND(REQ := FALSE,
                              LEN := #statSend.tsendFct.dataOffset,
                              ID := #tempConnOucId,
                              DATA := #statSend.tsendFct.data);

                   #instTRCV(EN_R := FALSE,
                             ID := #diagnostics.localConfig.connection.connectionID,
                             LEN := 0,
                             ADHOC := TRUE,
                             NDR => #statReceive.trcvFct.dataReceived,
                             RCVD_LEN => #statReceive.trcvFct.dataLength,
                             DATA := #statReceive.trcvFct.data);

                   #instTDISCON(REQ := TRUE,
                                ID := #tempConnOucId);

                   //Error occurred during processing
                   IF (#instTDISCON.ERROR) THEN

                       #statDiag.bufferIndex := #statDiag.bufferIndex + 1;
                       #statDiag.buffer[#statDiag.bufferIndex].status := #ERR_CLOSE_CONNECTION;
                       #statDiag.buffer[#statDiag.bufferIndex].subFunctionErrorID := #instTDISCON.STATUS;
                       #statDiag.buffer[#statDiag.bufferIndex].additionalValue1 := 0.0;
                       #statDiag.buffer[#statDiag.bufferIndex].additionalValue2 := 0.0;
                       #statDiag.buffer[#statDiag.bufferIndex].additionalValue3 := 0.0;
                       #statDiag.buffer[#statDiag.bufferIndex].additionalValue4 := T#0ms;

                       #statState.connection := #STATE_INACTIVE_PREPARE;

                       #instTDISCON(REQ := FALSE,
                                    ID := #tempConnOucId);

                   ELSIF (#instTDISCON.DONE) THEN

                       #instTDISCON(REQ := FALSE,
                                    ID := #tempConnOucId);
                       //Job executed without errors
                       IF (#enable AND (NOT #statFallingEdgeEnable)) THEN
                           //Reconnect automatically if not in disconnecting process
                           #statIterator := 0;
                           #statState.connection := #STATE_WAIT;
                       ELSE
                           //Reset all active failures in the diagnostics buffer
                           FOR #statIterator := 0 TO #DIAG_BUFFER_UPPER_LIM BY 1 DO
                               #diagnostics.buffer[#statIterator].isActive := FALSE;
                           END_FOR;

                           #statState.connection := #STATE_INACTIVE_PREPARE;
                       END_IF;
                       //Job is not completed yet
                   ELSE
                       ;//Wait until job is finished
                   END_IF;
               END_REGION CALL_TDISCON

           #ERROR_STATE:
               REGION ERROR
                   ;
               END_REGION ERROR
       END_CASE;
   END_REGION STATE_MACHINE

   REGION DIAGNOSTICS
       // -----------------------------------------------------------------------------------------------------------
       //Diagnostics buffer
       // -----------------------------------------------------------------------------------------------------------
   diag:
       //Diagnostics entry is in the temp. buffer
       IF (#statDiag.bufferIndex <> -1) THEN

           //Get current time
           #statRet := RD_LOC_T(#tempActTime);
           //init
           #statDiag.actualIndex := 0;

           WHILE (#statDiag.actualIndex <= #statDiag.bufferIndex) DO

               #tempUDint := 0;
               //Check if the failure is already in the buffer and still active
               FOR #statIterator := 0 TO #DIAG_BUFFER_UPPER_LIM BY 1 DO

                   IF (#diagnostics.buffer[#statIterator].isActive = TRUE) THEN

                       IF ((#statDiag.buffer[#statDiag.actualIndex].status = #WARN_SEND_CYCLE_EXPIRED)
                           AND
                           (#diagnostics.buffer[#statIterator].status = #WARN_SEND_CYCLE_EXPIRED)
                           AND
                           (#diagnostics.buffer[#statIterator].additionalValue1 = #statDiag.buffer[#statDiag.actualIndex].additionalValue1)
                           AND
                           (#diagnostics.buffer[#statIterator].additionalValue2 = #statDiag.buffer[#statDiag.actualIndex].additionalValue2)
                           AND
                           (#diagnostics.buffer[#statIterator].additionalValue3 = #statDiag.buffer[#statDiag.actualIndex].additionalValue3)) THEN
                           //Retrigger just the activation time
                           #diagnostics.buffer[#statIterator].timestamp := #tempActTime;
                           #diagnostics.buffer[#statIterator].additionalValue4 := #statDiag.buffer[#statDiag.actualIndex].additionalValue4;
                           #tempUDint := 100;
                           EXIT;
                       ELSIF ((#diagnostics.buffer[#statIterator].status = #statDiag.buffer[#statDiag.actualIndex].status)
                           AND
                           (#diagnostics.buffer[#statIterator].additionalValue1 = #statDiag.buffer[#statDiag.actualIndex].additionalValue1)
                           AND
                           (#diagnostics.buffer[#statIterator].additionalValue2 = #statDiag.buffer[#statDiag.actualIndex].additionalValue2)
                           AND
                           (#diagnostics.buffer[#statIterator].additionalValue3 = #statDiag.buffer[#statDiag.actualIndex].additionalValue3)
                           AND
                           (#diagnostics.buffer[#statIterator].additionalValue4 = #statDiag.buffer[#statDiag.actualIndex].additionalValue4)) THEN
                           //Retrigger just the activation time
                           #diagnostics.buffer[#statIterator].timestamp := #tempActTime;
                           #tempUDint := 100;
                           EXIT;
                       ELSE
                           ;//ErrorId is not in the diagnostics buffer
                       END_IF;
                   END_IF;
               END_FOR;

               IF (#tempUDint = 100) THEN
                   ;//ErrorId was already retriggered
               ELSE
                   //Check range of diagnostics ring buffer [0...DIAG_ARRAY]
                   IF ((#diagnostics.bufferIndex = 255) OR (#diagnostics.bufferIndex = #DIAG_BUFFER_UPPER_LIM)) THEN
                       #diagnostics.bufferIndex := 0;
                   ELSE
                       #diagnostics.bufferIndex := #diagnostics.bufferIndex + 1;
                   END_IF;

                   //Stored new entry in the diagnostics buffer
                   #diagnostics.buffer[#diagnostics.bufferIndex].status := #statDiag.buffer[#statDiag.actualIndex].status;
                   #diagnostics.buffer[#diagnostics.bufferIndex].timestamp := #tempActTime;
                   #diagnostics.buffer[#diagnostics.bufferIndex].isActive := TRUE;

                   #diagnostics.buffer[#diagnostics.bufferIndex].subFunctionErrorID := #statDiag.buffer[#statDiag.actualIndex].subFunctionErrorID;
                   #diagnostics.buffer[#diagnostics.bufferIndex].additionalValue1 := #statDiag.buffer[#statDiag.actualIndex].additionalValue1;
                   #diagnostics.buffer[#diagnostics.bufferIndex].additionalValue2 := #statDiag.buffer[#statDiag.actualIndex].additionalValue2;
                   #diagnostics.buffer[#diagnostics.bufferIndex].additionalValue3 := #statDiag.buffer[#statDiag.actualIndex].additionalValue3;
                   #diagnostics.buffer[#diagnostics.bufferIndex].additionalValue4 := #statDiag.buffer[#statDiag.actualIndex].additionalValue4;
               END_IF;

               IF ((#diagnostics.buffer[#diagnostics.bufferIndex].status = #STATUS_TCP_CONNECTED)
                   OR (#diagnostics.buffer[#diagnostics.bufferIndex].status = #STATUS_CONNECTED_V1)
                   OR (#diagnostics.buffer[#diagnostics.bufferIndex].status = #STATUS_CONNECTED_V2))
               THEN
                   #statConnectAttempts := 0;
                   #diagnostics.statistics.lastConnect := #tempActTime;
               END_IF;

               //Set FB status
               #status := #statStatus := #statDiag.buffer[#statDiag.actualIndex].status;

               //Check if FB.error has been set ?
               IF ((#statDiag.buffer[#statDiag.actualIndex].status >= #ERR_COM_SERVICE)//16#8200
                   AND
                   (#statDiag.buffer[#statDiag.actualIndex].status <= #ERR_WRONG_TELEGRAM_ID))//16#8614
               THEN

                   #error := TRUE;
                   #connected := #statConnected := FALSE;
                   #sending := #statSending := FALSE;
                   #dataReceived := #statDataReceived := FALSE;
                   #receivedDataLength := 0;

                   //Check if FB.busy has been set ?
                   IF ((#statDiag.buffer[#statDiag.actualIndex].status >= #ERR_OPEN_CLIENT)//16#8600
                       AND
                       (#statDiag.buffer[#statDiag.actualIndex].status <= #ERR_WRONG_TELEGRAM_ID))//16#8614
                   THEN
                       #busy := TRUE;
                   ELSE
                       #busy := FALSE;
                   END_IF;

                   EXIT;//Leave loop
               ELSE
                   ;
               END_IF;

               //Increase index
               #statDiag.actualIndex := #statDiag.actualIndex + 1;

           END_WHILE;
       ELSE
           ;//No failure
       END_IF;//End: Diagnostics buffer
   END_REGION DIAGNOSTICS
END_FUNCTION_BLOCK
